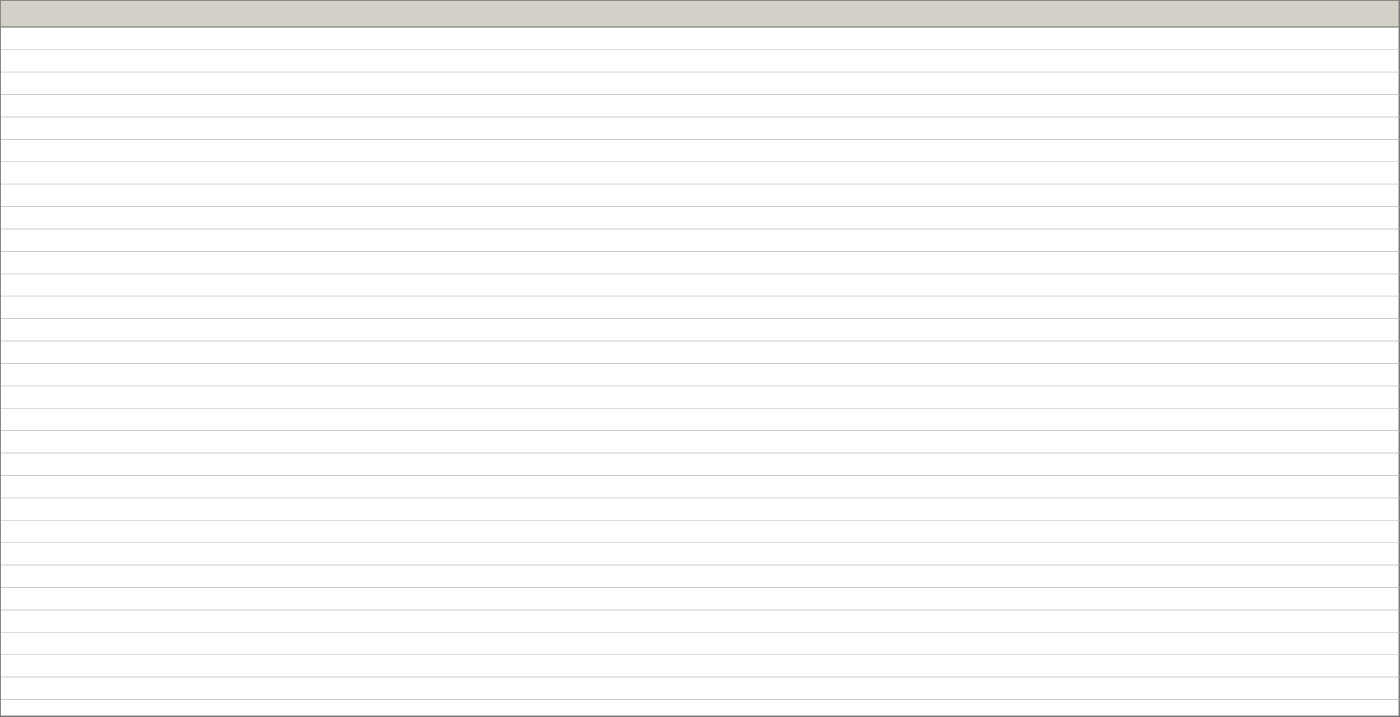
VISUALIZATION vis_Error_Search  // 1560x800
    Table (0,0 1560x800), data array: Buffer_Search_Messages
        p3854506369: Buffer_Search_Messages[INDEX].sDateTime
        p1892666644: Buffer_Search_Messages[INDEX].sErrID
        p338671338: Buffer_Search_Messages[INDEX].sLevel
        p2170511999: Buffer_Search_Messages[INDEX].sModuleDescription
        p3723444502: Buffer_Search_Messages[INDEX].sErrorMessage
        p4092479075: Module Description
        p2237128397: Error Message
END_VISUALIZATION

(* stored: Version 1.1.0.1, ProductVersion 3.1.4024.13
   Visu vis_Error_Search: Id {af0e7be7-8efe-4b7f-bdb4-cd7581603649} *)
